(* LS Electric XG5000 project: REMRES2 *)
(* PLC LSPLC *)

PROGRAM MainLD (* task: 스캔 프로그램 *)

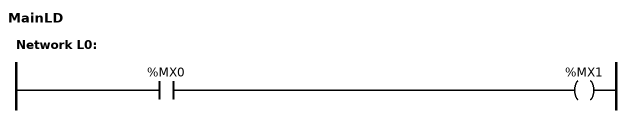
(* Rung L0 *)
%MX1 := %MX0;
END_PROGRAM

PROGRAM MainST (* task: 스캔 프로그램 *)
%MX1 := %MX0;
END_PROGRAM

PROGRAM MainIL (* task: 스캔 프로그램 *)
LD %MX0
ST %MX1
END_PROGRAM

PROGRAM MainSFC (* task: 스캔 프로그램 *)
VAR
    GOTO_INIT : BOOL;
    TRANS : BOOL;
END_VAR
(* SFC body not rendered *)
END_PROGRAM